FUNCTION_BLOCK fbMonostableRelay IMPLEMENTS iRelay
VAR
    RelayOutput AT %Q* : BOOL;
END_VAR

PROPERTY PUBLIC IsSet : BOOL
GET
IsSet := RelayOutput;
END_GET
END_PROPERTY

METHOD Reset
RelayOutput := FALSE;
END_METHOD

METHOD Set
RelayOutput := TRUE;
END_METHOD

END_FUNCTION_BLOCK

(* stored: Version 1.1.0.1
   POU fbMonostableRelay: Id {1e99fd58-1860-4d43-9df9-50b04eba5883}, SpecialFunc None
   Property IsSet: Id {01e1278e-4d38-47d2-93b5-d878fc42c631}
   Get Get: Id {df2cd450-f648-444f-8ba7-120d765e1ee5}
   Method Reset: Id {c8cf2292-1af8-451d-bc98-879376fef134}
   Method Set: Id {8b890796-e473-4154-bfe5-d2bb589f8e04} *)
